// TIA Portal V20 export
DATA_BLOCK "Melden_VisuAllgemein_DB"   // DB155
// stored: InstanceOfName Melden_VisuAllgemein, InstanceOfType FB
"Melden_VisuAllgemein"
   // VAR
   //    Register_leer : "Teile Status";
   //    auf_Seite_Richten { S7_SetPoint := 'True'} : Bool;
   //    Flanke_Bildwechsel { S7_SetPoint := 'True'} : R_TRIG;
   //    Bild_tmp { S7_SetPoint := 'True'} : DInt;
   //    WartezeitSicherung_Reset { S7_SetPoint := 'True'} : TON_TIME;
   //    Flanke_Türe8_schließen { S7_SetPoint := 'True'} : R_TRIG;
   //    Flanke_Türe8_öffnen { S7_SetPoint := 'True'} : R_TRIG;
   // END_VAR
   // VAR RETAIN
   //    Artikelnummer_tmp { ExternalAccessible := 'False'; ExternalVisible := 'False'; ExternalWritable := 'False'} : String;
   // END_VAR
   // VAR
   //    VZ_Leerfahren { S7_SetPoint := 'True'} : TON_TIME;
   // END_VAR
BEGIN
END_DATA_BLOCK
